            #Stored := "FRK_ConfigFind"(Scope := 'StationB.Satellite.Inner.Cell.Clamp', Key := 'preset', ModelCode := 'MODEL_A');
            IF #Stored > 0 THEN "FRK_ConfigStore".Rows[#Stored].Used := FALSE; END_IF;
            #Stored := "FRK_ConfigFind"(Scope := 'StationB.Satellite.Inner.Cell.Gate', Key := 'timeout', ModelCode := 'MODEL_A');
            IF #Stored > 0 THEN "FRK_ConfigStore".Rows[#Stored].Used := FALSE; END_IF;
            #Stored := "FRK_ConfigFind"(Scope := 'StationB.Satellite.Inner.Cell.Gate', Key := 'preset', ModelCode := 'MODEL_A');
            IF #Stored > 0 THEN "FRK_ConfigStore".Rows[#Stored].Used := FALSE; END_IF;
            "FRK_ConfigLoss"(RootIndex := 2, Scope := 'StationB');
        11:
            #Stored := "FRK_ConfigFind"(Scope := 'StationB', Key := 'timeout', ModelCode := 'MODEL_B');
            IF #Stored > 0 THEN "FRK_ConfigStore".Rows[#Stored].Used := FALSE; END_IF;
            #Stored := "FRK_ConfigFind"(Scope := 'StationB', Key := 'preset', ModelCode := 'MODEL_B');
            IF #Stored > 0 THEN "FRK_ConfigStore".Rows[#Stored].Used := FALSE; END_IF;
            #Stored := "FRK_ConfigFind"(Scope := 'StationB.Cell', Key := 'timeout', ModelCode := 'MODEL_B');
            IF #Stored > 0 THEN "FRK_ConfigStore".Rows[#Stored].Used := FALSE; END_IF;
            #Stored := "FRK_ConfigFind"(Scope := 'StationB.Cell', Key := 'preset', ModelCode := 'MODEL_B');
            IF #Stored > 0 THEN "FRK_ConfigStore".Rows[#Stored].Used := FALSE; END_IF;
            #Stored := "FRK_ConfigFind"(Scope := 'StationB.Cell.Clamp', Key := 'timeout', ModelCode := 'MODEL_B');
            IF #Stored > 0 THEN "FRK_ConfigStore".Rows[#Stored].Used := FALSE; END_IF;
            #Stored := "FRK_ConfigFind"(Scope := 'StationB.Cell.Clamp', Key := 'preset', ModelCode := 'MODEL_B');
            IF #Stored > 0 THEN "FRK_ConfigStore".Rows[#Stored].Used := FALSE; END_IF;
            #Stored := "FRK_ConfigFind"(Scope := 'StationB.Cell.Gate', Key := 'timeout', ModelCode := 'MODEL_B');
            IF #Stored > 0 THEN "FRK_ConfigStore".Rows[#Stored].Used := FALSE; END_IF;
            #Stored := "FRK_ConfigFind"(Scope := 'StationB.Cell.Gate', Key := 'preset', ModelCode := 'MODEL_B');
            IF #Stored > 0 THEN "FRK_ConfigStore".Rows[#Stored].Used := FALSE; END_IF;
            #Stored := "FRK_ConfigFind"(Scope := 'StationB.Satellite', Key := 'timeout', ModelCode := 'MODEL_B');
            IF #Stored > 0 THEN "FRK_ConfigStore".Rows[#Stored].Used := FALSE; END_IF;
            #Stored := "FRK_ConfigFind"(Scope := 'StationB.Satellite', Key := 'preset', ModelCode := 'MODEL_B');
            IF #Stored > 0 THEN "FRK_ConfigStore".Rows[#Stored].Used := FALSE; END_IF;
            #Stored := "FRK_ConfigFind"(Scope := 'StationB.Satellite.Cell', Key := 'timeout', ModelCode := 'MODEL_B');
            IF #Stored > 0 THEN "FRK_ConfigStore".Rows[#Stored].Used := FALSE; END_IF;
            #Stored := "FRK_ConfigFind"(Scope := 'StationB.Satellite.Cell', Key := 'preset', ModelCode := 'MODEL_B');
            IF #Stored > 0 THEN "FRK_ConfigStore".Rows[#Stored].Used := FALSE; END_IF;
            #Stored := "FRK_ConfigFind"(Scope := 'StationB.Satellite.Cell.Clamp', Key := 'timeout', ModelCode := 'MODEL_B');
            IF #Stored > 0 THEN "FRK_ConfigStore".Rows[#Stored].Used := FALSE; END_IF;
            #Stored := "FRK_ConfigFind"(Scope := 'StationB.Satellite.Cell.Clamp', Key := 'preset', ModelCode := 'MODEL_B');
            IF #Stored > 0 THEN "FRK_ConfigStore".Rows[#Stored].Used := FALSE; END_IF;
            #Stored := "FRK_ConfigFind"(Scope := 'StationB.Satellite.Cell.Gate', Key := 'timeout', ModelCode := 'MODEL_B');
            IF #Stored > 0 THEN "FRK_ConfigStore".Rows[#Stored].Used := FALSE; END_IF;
            #Stored := "FRK_ConfigFind"(Scope := 'StationB.Satellite.Cell.Gate', Key := 'preset', ModelCode := 'MODEL_B');
            IF #Stored > 0 THEN "FRK_ConfigStore".Rows[#Stored].Used := FALSE; END_IF;
            #Stored := "FRK_ConfigFind"(Scope := 'StationB.Satellite.Inner', Key := 'timeout', ModelCode := 'MODEL_B');
            IF #Stored > 0 THEN "FRK_ConfigStore".Rows[#Stored].Used := FALSE; END_IF;
            #Stored := "FRK_ConfigFind"(Scope := 'StationB.Satellite.Inner', Key := 'preset', ModelCode := 'MODEL_B');
            IF #Stored > 0 THEN "FRK_ConfigStore".Rows[#Stored].Used := FALSE; END_IF;
            #Stored := "FRK_ConfigFind"(Scope := 'StationB.Satellite.Inner.Cell', Key := 'timeout', ModelCode := 'MODEL_B');
            IF #Stored > 0 THEN "FRK_ConfigStore".Rows[#Stored].Used := FALSE; END_IF;
            #Stored := "FRK_ConfigFind"(Scope := 'StationB.Satellite.Inner.Cell', Key := 'preset', ModelCode := 'MODEL_B');
            IF #Stored > 0 THEN "FRK_ConfigStore".Rows[#Stored].Used := FALSE; END_IF;
            #Stored := "FRK_ConfigFind"(Scope := 'StationB.Satellite.Inner.Cell.Clamp', Key := 'timeout', ModelCode := 'MODEL_B');
            IF #Stored > 0 THEN "FRK_ConfigStore".Rows[#Stored].Used := FALSE; END_IF;
            #Stored := "FRK_ConfigFind"(Scope := 'StationB.Satellite.Inner.Cell.Clamp', Key := 'preset', ModelCode := 'MODEL_B');
            IF #Stored > 0 THEN "FRK_ConfigStore".Rows[#Stored].Used := FALSE; END_IF;
            #Stored := "FRK_ConfigFind"(Scope := 'StationB.Satellite.Inner.Cell.Gate', Key := 'timeout', ModelCode := 'MODEL_B');
            IF #Stored > 0 THEN "FRK_ConfigStore".Rows[#Stored].Used := FALSE; END_IF;
            #Stored := "FRK_ConfigFind"(Scope := 'StationB.Satellite.Inner.Cell.Gate', Key := 'preset', ModelCode := 'MODEL_B');
            IF #Stored > 0 THEN "FRK_ConfigStore".Rows[#Stored].Used := FALSE; END_IF;
            "FRK_ConfigLoss"(RootIndex := 2, Scope := 'StationB');
        12:
            "FRK_AccessPolicies".Rows[2].Scope := 'StationB';
            "FRK_AccessPolicies".Rows[2].SchemaVersion := 0;
            "FRK_AccessPolicies".Rows[2].Initialized := TRUE;
        13:
            "FRK_SetStore".Sets[2, 1].Info.Used := FALSE;
            "FRK_ConfigLoss"(RootIndex := 2, Scope := 'StationB');
        14:
            "FRK_SetStore".Sets[2, 2].Info.Used := FALSE;
            "FRK_ConfigLoss"(RootIndex := 2, Scope := 'StationB');
        15:
            "FRK_SetStore".Sets[2, 3].Info.Used := FALSE;
            "FRK_ConfigLoss"(RootIndex := 2, Scope := 'StationB');
        16:
            "FRK_SetStore".Sets[2, 4].Info.Used := FALSE;
            "FRK_ConfigLoss"(RootIndex := 2, Scope := 'StationB');
        17:
            "FRK_LocalUsers".SchemaVersion := 0; "FRK_LocalUsers".Generation := 0; "FRK_LocalUsers".Checksum := DWORD#0;
            "FRK_AccessStorage".UsersCommissioned := TRUE; "FRK_AccessStorage".UsersReady := FALSE; "FRK_AccessStorage".UsersLost := TRUE;
        ELSE RETURN;
    END_CASE;
END_FUNCTION
FUNCTION "FRK_DocCapture" : Void
{ S7_Optimized_Access := 'TRUE' }
VERSION : 0.1
VAR_INPUT
    Slot : Int;
END_VAR
VAR_IN_OUT
    Ok : Bool;
    Length : DInt;
END_VAR
BEGIN
    #Ok := FALSE; #Length := 0;
    CASE #Slot OF
        1: #Ok := "FRK_DocCapture_D001"(Length := #Length);
        2: #Ok := "FRK_DocCapture_D002"(Length := #Length);
        3: #Ok := "FRK_DocCapture_D003"(Length := #Length);
        4: #Ok := "FRK_DocCapture_D004"(Length := #Length);
        5: #Ok := "FRK_DocCapture_D005"(Length := #Length);
        6: #Ok := "FRK_DocCapture_D006"(Length := #Length);
        7: #Ok := "FRK_DocCapture_D007"(Length := #Length);
        8: #Ok := "FRK_DocCapture_D008"(Length := #Length);
        9: #Ok := "FRK_DocCapture_D009"(Length := #Length);
        10: #Ok := "FRK_DocCapture_D010"(Length := #Length);
        11: #Ok := "FRK_DocCapture_D011"(Length := #Length);
        12: #Ok := "FRK_DocCapture_D012"(Length := #Length);
        13: #Ok := "FRK_DocCapture_D013"(Length := #Length);
        14: #Ok := "FRK_DocCapture_D014"(Length := #Length);
        15: #Ok := "FRK_DocCapture_D015"(Length := #Length);
        16: #Ok := "FRK_DocCapture_D016"(Length := #Length);
        17: #Ok := "FRK_DocCapture_D017"(Length := #Length);
        ELSE RETURN;
    END_CASE;
END_FUNCTION
FUNCTION "FRK_DocApply" : Bool
{ S7_Optimized_Access := 'TRUE' }
VERSION : 0.1
VAR_INPUT
    Slot : Int;
END_VAR
BEGIN
    #FRK_DocApply := FALSE;
    CASE #Slot OF
        1: #FRK_DocApply := "FRK_DocApply_D001"();
        2: #FRK_DocApply := "FRK_DocApply_D002"();
        3: #FRK_DocApply := "FRK_DocApply_D003"();
        4: #FRK_DocApply := "FRK_DocApply_D004"();
        5: #FRK_DocApply := "FRK_DocApply_D005"();
        6: #FRK_DocApply := "FRK_DocApply_D006"();
        7: #FRK_DocApply := "FRK_DocApply_D007"();
        8: #FRK_DocApply := "FRK_DocApply_D008"();
        9: #FRK_DocApply := "FRK_DocApply_D009"();
        10: #FRK_DocApply := "FRK_DocApply_D010"();
        11: #FRK_DocApply := "FRK_DocApply_D011"();
        12: #FRK_DocApply := "FRK_DocApply_D012"();
        13: #FRK_DocApply := "FRK_DocApply_D013"();
        14: #FRK_DocApply := "FRK_DocApply_D014"();
        15: #FRK_DocApply := "FRK_DocApply_D015"();
        16: #FRK_DocApply := "FRK_DocApply_D016"();
        17: #FRK_DocApply := "FRK_DocApply_D017"();
        ELSE RETURN;
    END_CASE;
END_FUNCTION
FUNCTION "FRK_DocBoot" : Void
{ S7_Optimized_Access := 'TRUE' }
VERSION : 0.1
VAR_INPUT
    Startup : Bool;
END_VAR
VAR_IN_OUT
    Ready : Bool;
END_VAR
VAR_TEMP
    Slot : Int;
    Done : Bool;
    Ok : Bool;
END_VAR
BEGIN
    IF #Startup THEN
        "FRK_PersistConsumers".Ready := FALSE;
        FOR #Slot := 1 TO 17 DO
            "FRK_PersistConsumers".Rows[#Slot].State := 0; "FRK_PersistConsumers".Rows[#Slot].Ticket := 0;
            "FRK_PersistConsumers".Rows[#Slot].Dirty := FALSE; "FRK_PersistConsumers".Rows[#Slot].Failed := FALSE;
            "FRK_PersistConsumers".Rows[#Slot].Rejected := FALSE; "FRK_PersistConsumers".Rows[#Slot].Acknowledged := FALSE;
            "FRK_PersistConsumers".Rows[#Slot].RetrySince := "FRK_Clock".NowMs;
            "FRK_PersistConsumers".Rows[#Slot].PendingSince := LDT#1970-01-01-00:00:00;
            "FRK_PersistConsumers".Rows[#Slot].NextSince := LDT#1970-01-01-00:00:00;
        END_FOR;
    END_IF;
    #Ready := TRUE;
    "FRK_PersistStatus".Failed := FALSE;
    FOR #Slot := 1 TO 17 DO
        IF "FRK_PersistConsumers".Rows[#Slot].State = 0 THEN
            IF NOT "FRK_PersistConsumers".Rows[#Slot].Failed OR "FRK_Elapsed"(NewMs := "FRK_Clock".NowMs, OldMs := "FRK_PersistConsumers".Rows[#Slot].RetrySince) >= 1000 THEN
                "FRK_PersistConsumers".Rows[#Slot].Ticket := "FRK_PersistStart"(Slot := #Slot, WriteDocument := FALSE, Length := 0);
                IF "FRK_PersistConsumers".Rows[#Slot].Ticket <> 0 THEN "FRK_PersistConsumers".Rows[#Slot].State := 1; END_IF;
            END_IF;
        ELSIF "FRK_PersistConsumers".Rows[#Slot].State = 1 THEN
            #Done := "FRK_PersistPoll"(Ticket := "FRK_PersistConsumers".Rows[#Slot].Ticket, Result := "FRK_PersistConsumers".Rows[#Slot].Result);
            IF #Done THEN
                "FRK_PersistConsumers".Rows[#Slot].Ticket := 0;
                IF NOT "FRK_PersistConsumers".Rows[#Slot].Result.Ok THEN
                    "FRK_PersistConsumers".Rows[#Slot].Failed := TRUE; "FRK_PersistConsumers".Rows[#Slot].State := 0;
                    "FRK_PersistConsumers".Rows[#Slot].RetrySince := "FRK_Clock".NowMs;
                ELSE
                    "FRK_PersistConsumers".Rows[#Slot].Failed := FALSE;
                    #Ok := NOT "FRK_PersistConsumers".Rows[#Slot].Result.Lost;
                    "FRK_PersistConsumers".Rows[#Slot].Virgin := #Ok AND NOT "FRK_PersistConsumers".Rows[#Slot].Result.Found;
                    IF #Ok AND "FRK_PersistConsumers".Rows[#Slot].Result.Found THEN #Ok := "FRK_DocApply"(Slot := #Slot); END_IF;
                    IF NOT #Ok THEN
                        "FRK_DocReject"(Slot := #Slot);
                        "FRK_PersistConsumers".Rows[#Slot].Rejected := TRUE;
                    ELSIF "FRK_PersistConsumers".Rows[#Slot].Virgin THEN "FRK_PersistDirty"(Slot := #Slot); END_IF;
                    "FRK_PersistConsumers".Rows[#Slot].State := 2;
                END_IF;
            END_IF;
        END_IF;
        IF "FRK_PersistConsumers".Rows[#Slot].State <> 2 THEN #Ready := FALSE; END_IF;
        "FRK_PersistStatus".Failed := "FRK_PersistStatus".Failed OR "FRK_PersistConsumers".Rows[#Slot].Failed;
    END_FOR;
    "FRK_PersistStatus".Restoring := NOT #Ready;
    "FRK_PersistStatus".NativeStatus := INT_TO_WORD("FRK_PersistRuntime".NativeResult);
    "FRK_PersistConsumers".Ready := #Ready;
END_FUNCTION
FUNCTION "FRK_DocCyclic" : Void
{ S7_Optimized_Access := 'TRUE' }
VERSION : 0.1
VAR_TEMP
    Slot : Int;
    Done : Bool;
    Ok : Bool;
    Length : DInt;
END_VAR
BEGIN
    IF NOT "FRK_PersistConsumers".Ready THEN RETURN; END_IF;
    FOR #Slot := 1 TO 17 DO
        IF "FRK_PersistConsumers".Rows[#Slot].Ticket <> 0 THEN
            #Done := "FRK_PersistPoll"(Ticket := "FRK_PersistConsumers".Rows[#Slot].Ticket, Result := "FRK_PersistConsumers".Rows[#Slot].Result);
            IF #Done THEN
                "FRK_PersistConsumers".Rows[#Slot].Ticket := 0;
                "FRK_PersistConsumers".Rows[#Slot].Failed := NOT "FRK_PersistConsumers".Rows[#Slot].Result.Ok;
                "FRK_PersistConsumers".Rows[#Slot].RetrySince := "FRK_Clock".NowMs;
                IF "FRK_PersistConsumers".Rows[#Slot].Failed THEN "FRK_PersistConsumers".Rows[#Slot].Dirty := TRUE;
                ELSIF "FRK_PersistConsumers".Rows[#Slot].Dirty THEN "FRK_PersistConsumers".Rows[#Slot].PendingSince := "FRK_PersistConsumers".Rows[#Slot].NextSince;
                ELSE "FRK_PersistConsumers".Rows[#Slot].PendingSince := LDT#1970-01-01-00:00:00; END_IF;
            END_IF;
        ELSIF "FRK_PersistConsumers".Rows[#Slot].Dirty AND (NOT "FRK_PersistConsumers".Rows[#Slot].Rejected OR "FRK_PersistConsumers".Rows[#Slot].Acknowledged) THEN
            IF NOT "FRK_PersistConsumers".Rows[#Slot].Failed OR "FRK_Elapsed"(NewMs := "FRK_Clock".NowMs, OldMs := "FRK_PersistConsumers".Rows[#Slot].RetrySince) >= 1000 THEN
                "FRK_DocCapture"(Slot := #Slot, Ok := #Ok, Length := #Length);
                IF #Ok THEN
                    "FRK_PersistConsumers".Rows[#Slot].Ticket := "FRK_PersistStart"(Slot := #Slot, WriteDocument := TRUE, Length := #Length);
                    IF "FRK_PersistConsumers".Rows[#Slot].Ticket <> 0 THEN "FRK_PersistConsumers".Rows[#Slot].Dirty := FALSE; END_IF;
                ELSE "FRK_PersistConsumers".Rows[#Slot].Failed := TRUE; "FRK_PersistConsumers".Rows[#Slot].RetrySince := "FRK_Clock".NowMs; END_IF;
            END_IF;
        END_IF;
    END_FOR;
END_FUNCTION
